FUNCTION_BLOCK CASE_SEQUENCER (* Migrated from IEC 61131-3 ST *)
  (* Standard: 61499-2 *)
  (* Version 1.0, 2026-11-06, st2fb *)
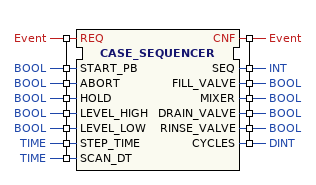
  EVENT_INPUT
    REQ WITH START_PB, ABORT, HOLD, LEVEL_HIGH, LEVEL_LOW, STEP_TIME, SCAN_DT;
  END_EVENT
  EVENT_OUTPUT
    CNF WITH SEQ, FILL_VALVE, MIXER, DRAIN_VALVE, RINSE_VALVE, CYCLES;
  END_EVENT
  VAR_INPUT
    START_PB : BOOL;
    ABORT : BOOL;
    HOLD : BOOL;
    LEVEL_HIGH : BOOL;
    LEVEL_LOW : BOOL;
    STEP_TIME : TIME;
    SCAN_DT : TIME;
  END_VAR
  VAR_OUTPUT
    SEQ : INT;
    FILL_VALVE : BOOL;
    MIXER : BOOL;
    DRAIN_VALVE : BOOL;
    RINSE_VALVE : BOOL;
    CYCLES : DINT;
  END_VAR
  VAR
    TIMING : BOOL := FALSE;
    STEP_TIMER_IN : BOOL := FALSE;
    STEP_TIMER_PT : TIME := T#0s;
    STEP_TIMER_Q : BOOL := FALSE;
    STEP_TIMER_ET : TIME := T#0s;
    STEP_TIMER_STATE : INT := 0;
    STEP_TIMER_PREV_IN : BOOL := FALSE;
    STEP_TIMER_START_TIME : TIME := T#0s;
    ST2FB_NOW : TIME := T#0s;
  END_VAR
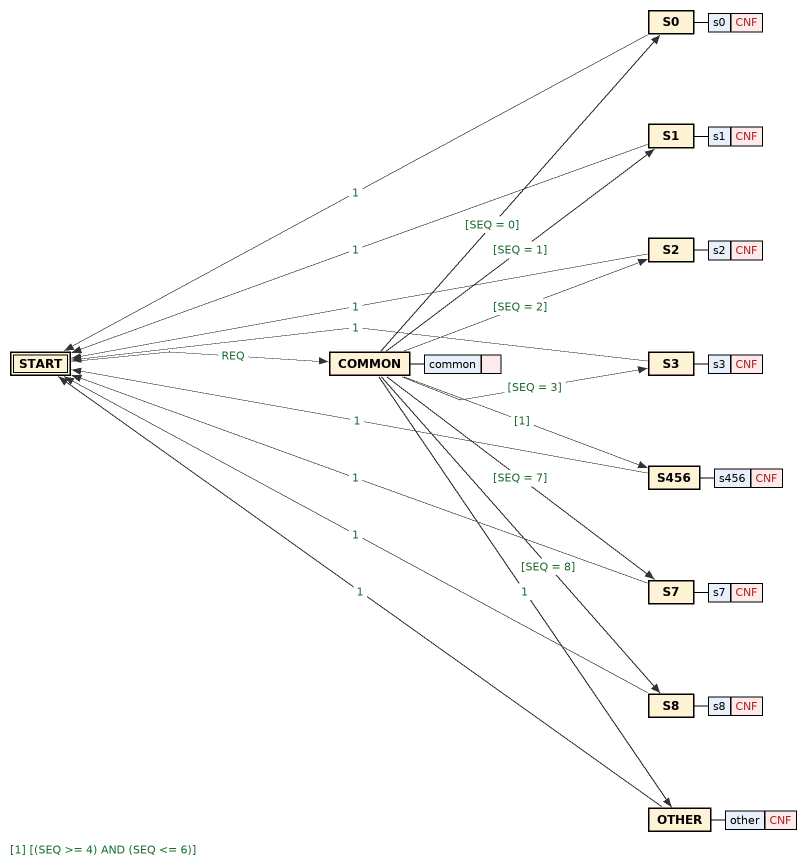
  EC_STATES
    START;
    COMMON : common;
    S0 : s0 -> CNF;
    S1 : s1 -> CNF;
    S2 : s2 -> CNF;
    S3 : s3 -> CNF;
    S456 : s456 -> CNF;
    S7 : s7 -> CNF;
    S8 : s8 -> CNF;
    OTHER : other -> CNF;
  END_STATES
  EC_TRANSITIONS
    START TO COMMON := REQ;
    COMMON TO S0 := [SEQ = 0];
    COMMON TO S1 := [SEQ = 1];
    COMMON TO S2 := [SEQ = 2];
    COMMON TO S3 := [SEQ = 3];
    COMMON TO S456 := [(SEQ >= 4) AND (SEQ <= 6)];
    COMMON TO S7 := [SEQ = 7];
    COMMON TO S8 := [SEQ = 8];
    COMMON TO OTHER := 1;
    S0 TO START := 1;
    S1 TO START := 1;
    S2 TO START := 1;
    S3 TO START := 1;
    S456 TO START := 1;
    S7 TO START := 1;
    S8 TO START := 1;
    OTHER TO START := 1;
  END_TRANSITIONS
  ALGORITHM common IN ST:
ST2FB_NOW := ST2FB_NOW + SCAN_DT;
IF NOT HOLD THEN
  STEP_TIMER_IN := TIMING;
  STEP_TIMER_PT := STEP_TIME;
  IF (STEP_TIMER_STATE = 0) AND NOT STEP_TIMER_PREV_IN AND STEP_TIMER_IN THEN
    STEP_TIMER_STATE := 1;
    STEP_TIMER_Q := FALSE;
    STEP_TIMER_START_TIME := ST2FB_NOW;
  ELSE
    IF NOT STEP_TIMER_IN THEN
      STEP_TIMER_ET := T#0s;
      STEP_TIMER_Q := FALSE;
      STEP_TIMER_STATE := 0;
    ELSIF STEP_TIMER_STATE = 1 THEN
      IF STEP_TIMER_START_TIME + STEP_TIMER_PT <= ST2FB_NOW THEN
        STEP_TIMER_STATE := 2;
        STEP_TIMER_Q := TRUE;
        STEP_TIMER_ET := STEP_TIMER_PT;
      ELSE
        STEP_TIMER_ET := ST2FB_NOW - STEP_TIMER_START_TIME;
      END_IF;
    END_IF;
  END_IF;
  STEP_TIMER_PREV_IN := STEP_TIMER_IN;
END_IF;
FILL_VALVE := FALSE;
MIXER := FALSE;
DRAIN_VALVE := FALSE;
RINSE_VALVE := FALSE;
IF ABORT THEN
  SEQ := 8;
END_IF;
  END_ALGORITHM
  ALGORITHM s0 IN ST:
TIMING := FALSE;
IF START_PB THEN
  SEQ := 1;
END_IF;
  END_ALGORITHM
  ALGORITHM s1 IN ST:
FILL_VALVE := TRUE;
IF LEVEL_HIGH THEN
  SEQ := 2;
  TIMING := TRUE;
END_IF;
  END_ALGORITHM
  ALGORITHM s2 IN ST:
MIXER := TRUE;
IF STEP_TIMER_Q THEN
  SEQ := 3;
  TIMING := FALSE;
END_IF;
  END_ALGORITHM
  ALGORITHM s3 IN ST:
DRAIN_VALVE := TRUE;
IF LEVEL_LOW THEN
  SEQ := 4;
END_IF;
  END_ALGORITHM
  ALGORITHM s456 IN ST:
RINSE_VALVE := TRUE;
IF STEP_TIMER_Q THEN
  SEQ := SEQ + 1;
  TIMING := FALSE;
ELSE
  TIMING := TRUE;
END_IF;
  END_ALGORITHM
  ALGORITHM s7 IN ST:
CYCLES := CYCLES + 1;
SEQ := 0;
  END_ALGORITHM
  ALGORITHM s8 IN ST:
TIMING := FALSE;
DRAIN_VALVE := TRUE;
IF LEVEL_LOW AND NOT ABORT THEN
  SEQ := 0;
END_IF;
  END_ALGORITHM
  ALGORITHM other IN ST:
SEQ := 0;
  END_ALGORITHM
END_FUNCTION_BLOCK
